(* Logix 5000 project; controller NWGG_Treater_Dayton vendor 1 type 14 code 238 rev 35.11; software revision 35.00; part 4 of 5 *)
(* tags used below, declared in another part *)
   Auto_Start_Treater : BOOL;
   Chemicals_Required : BOOL;
   Clear_Treater_Fault : BOOL;
   Current_Treater_Speed_Percent : REAL;
   Grain_Rate_CWT : REAL;
   IDX : DINT;
   K_Valve_ACK : BOOL;
   Manual_Start_Treater : BOOL;
   Non_Water_Total_Chemical_Package : REAL;
   Non_Water_Treatment_Package : REAL;
   SAIZeroScale : SAI_Zero_Scale[30];
   Start_Treating : BOOL;
   Stop_Treater : BOOL;
   tmrStartTreat : TIMER;
   tmrStopTreat : TIMER;
   Total_Chemical_Package : REAL;
   Treater_Pump : Treater_Pump[50];
   Treater_Running : BOOL;
   Treater_Speed_Percent : REAL;
   Water : Analog_Gallon_Values;
   Water_Control : Water_Pump_Control;
(* MainProgram, continued *)

ROUTINE Set_Scale_Values   (* ladder *)
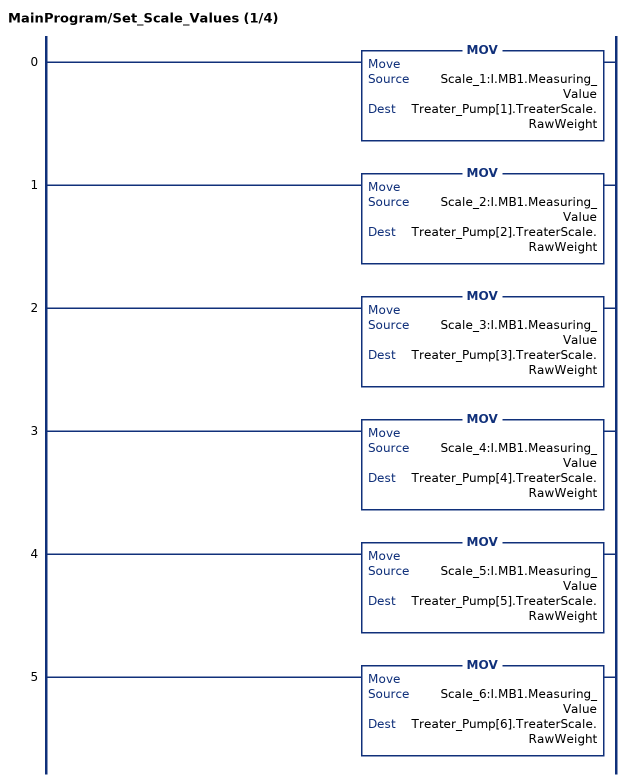
   0: MOV(Scale_1:I.MB1.Measuring_Value,Treater_Pump[1].TreaterScale.RawWeight);
   1: MOV(Scale_2:I.MB1.Measuring_Value,Treater_Pump[2].TreaterScale.RawWeight);
   2: MOV(Scale_3:I.MB1.Measuring_Value,Treater_Pump[3].TreaterScale.RawWeight);
   3: MOV(Scale_4:I.MB1.Measuring_Value,Treater_Pump[4].TreaterScale.RawWeight);
   4: MOV(Scale_5:I.MB1.Measuring_Value,Treater_Pump[5].TreaterScale.RawWeight);
   5: MOV(Scale_6:I.MB1.Measuring_Value,Treater_Pump[6].TreaterScale.RawWeight);
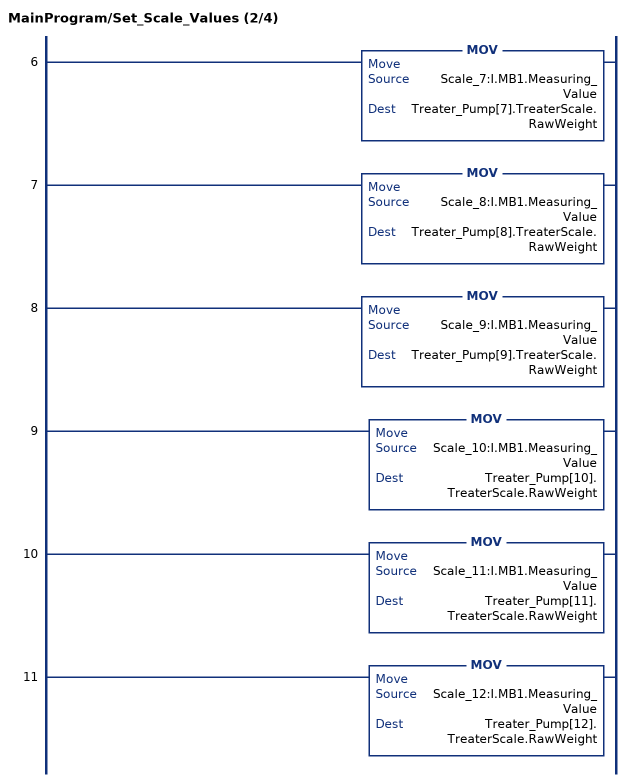
   6: MOV(Scale_7:I.MB1.Measuring_Value,Treater_Pump[7].TreaterScale.RawWeight);
   7: MOV(Scale_8:I.MB1.Measuring_Value,Treater_Pump[8].TreaterScale.RawWeight);
   8: MOV(Scale_9:I.MB1.Measuring_Value,Treater_Pump[9].TreaterScale.RawWeight);
   9: MOV(Scale_10:I.MB1.Measuring_Value,Treater_Pump[10].TreaterScale.RawWeight);
   10: MOV(Scale_11:I.MB1.Measuring_Value,Treater_Pump[11].TreaterScale.RawWeight);
   11: MOV(Scale_12:I.MB1.Measuring_Value,Treater_Pump[12].TreaterScale.RawWeight);
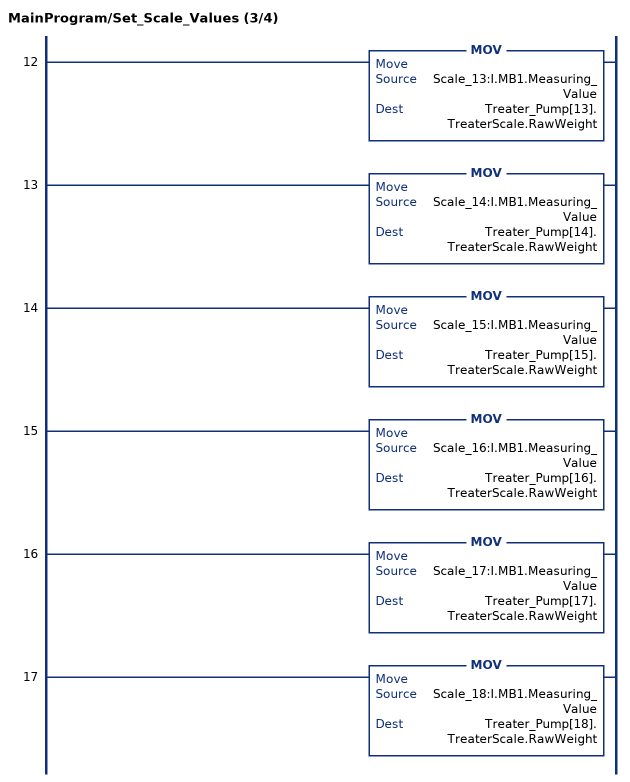
   12: MOV(Scale_13:I.MB1.Measuring_Value,Treater_Pump[13].TreaterScale.RawWeight);
   13: MOV(Scale_14:I.MB1.Measuring_Value,Treater_Pump[14].TreaterScale.RawWeight);
   14: MOV(Scale_15:I.MB1.Measuring_Value,Treater_Pump[15].TreaterScale.RawWeight);
   15: MOV(Scale_16:I.MB1.Measuring_Value,Treater_Pump[16].TreaterScale.RawWeight);
   16: MOV(Scale_17:I.MB1.Measuring_Value,Treater_Pump[17].TreaterScale.RawWeight);
   17: MOV(Scale_18:I.MB1.Measuring_Value,Treater_Pump[18].TreaterScale.RawWeight);
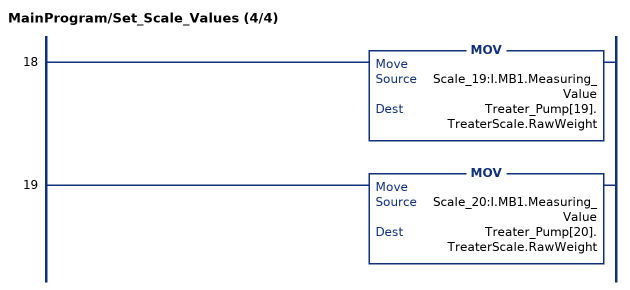
   18: MOV(Scale_19:I.MB1.Measuring_Value,Treater_Pump[19].TreaterScale.RawWeight);
   19: MOV(Scale_20:I.MB1.Measuring_Value,Treater_Pump[20].TreaterScale.RawWeight);
END_ROUTINE

ROUTINE SetHMIArrayIndex   (* ladder *)
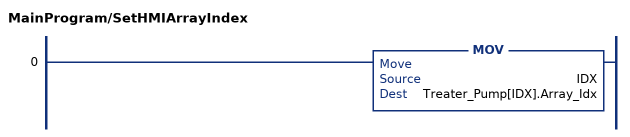
   0: MOV(IDX,Treater_Pump[IDX].Array_Idx);
END_ROUTINE

ROUTINE Treater   (* ladder *)
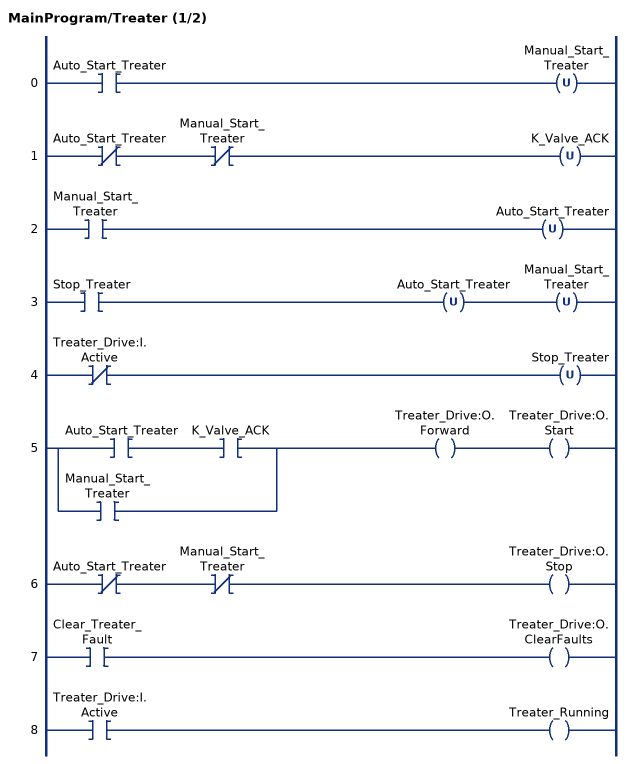
   0: XIC(Auto_Start_Treater)OTU(Manual_Start_Treater);
   1: XIO(Auto_Start_Treater)XIO(Manual_Start_Treater)OTU(K_Valve_ACK);
   2: XIC(Manual_Start_Treater)OTU(Auto_Start_Treater);
   3: XIC(Stop_Treater)OTU(Auto_Start_Treater)OTU(Manual_Start_Treater);
   4: XIO(Treater_Drive:I.Active)OTU(Stop_Treater);
   5: [XIC(Auto_Start_Treater) XIC(K_Valve_ACK) ,XIC(Manual_Start_Treater) ]OTE(Treater_Drive:O.Forward)OTE(Treater_Drive:O.Start);
   6: XIO(Auto_Start_Treater)XIO(Manual_Start_Treater)OTE(Treater_Drive:O.Stop);
   7: XIC(Clear_Treater_Fault)OTE(Treater_Drive:O.ClearFaults);
   8: XIC(Treater_Drive:I.Active)OTE(Treater_Running);
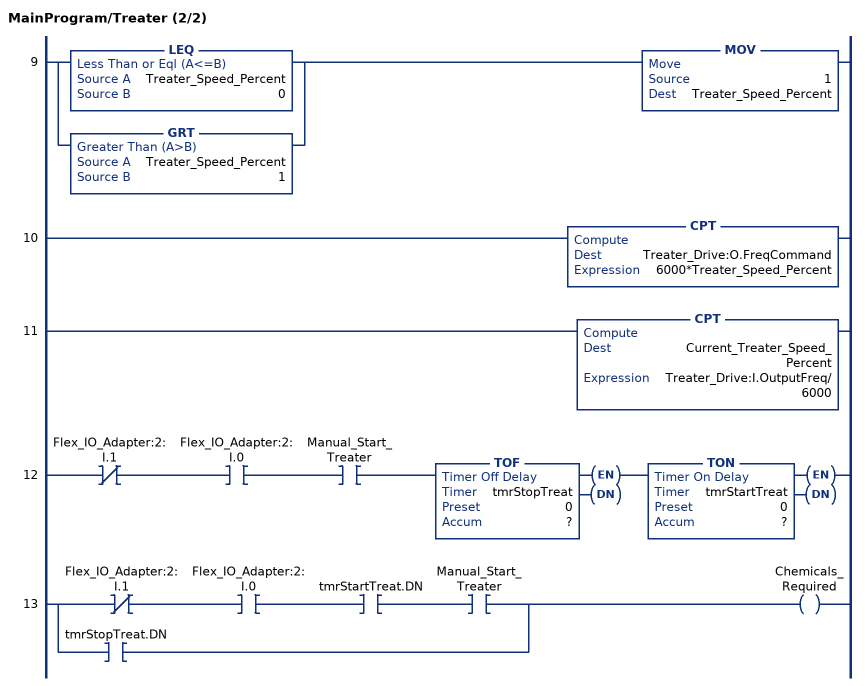
   9: [LEQ(Treater_Speed_Percent,0) ,GRT(Treater_Speed_Percent,1) ]MOV(1,Treater_Speed_Percent);
   10: CPT(Treater_Drive:O.FreqCommand,6000*Treater_Speed_Percent);
   11: CPT(Current_Treater_Speed_Percent,Treater_Drive:I.OutputFreq/6000);
   12: XIO(Flex_IO_Adapter:2:I.1)XIC(Flex_IO_Adapter:2:I.0)XIC(Manual_Start_Treater)TOF(tmrStopTreat,?,?)TON(tmrStartTreat,?,?);
   13: [XIO(Flex_IO_Adapter:2:I.1) XIC(Flex_IO_Adapter:2:I.0) XIC(tmrStartTreat.DN) XIC(Manual_Start_Treater) ,XIC(tmrStopTreat.DN) ]OTE(Chemicals_Required);
END_ROUTINE

ROUTINE Zero_Scales   (* ladder *)
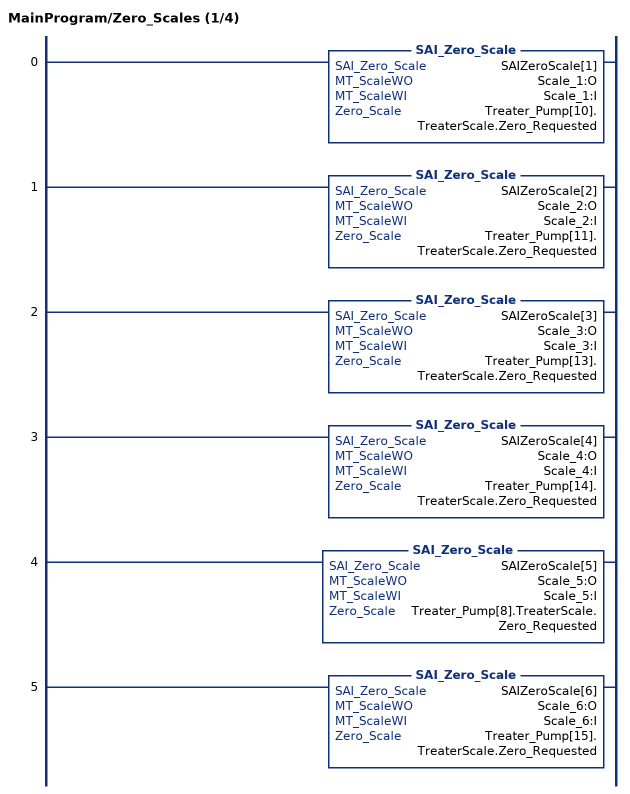
   0: SAI_Zero_Scale(SAIZeroScale[1],Scale_1:O,Scale_1:I,Treater_Pump[10].TreaterScale.Zero_Requested);
   1: SAI_Zero_Scale(SAIZeroScale[2],Scale_2:O,Scale_2:I,Treater_Pump[11].TreaterScale.Zero_Requested);
   2: SAI_Zero_Scale(SAIZeroScale[3],Scale_3:O,Scale_3:I,Treater_Pump[13].TreaterScale.Zero_Requested);
   3: SAI_Zero_Scale(SAIZeroScale[4],Scale_4:O,Scale_4:I,Treater_Pump[14].TreaterScale.Zero_Requested);
   4: SAI_Zero_Scale(SAIZeroScale[5],Scale_5:O,Scale_5:I,Treater_Pump[8].TreaterScale.Zero_Requested);
   5: SAI_Zero_Scale(SAIZeroScale[6],Scale_6:O,Scale_6:I,Treater_Pump[15].TreaterScale.Zero_Requested);
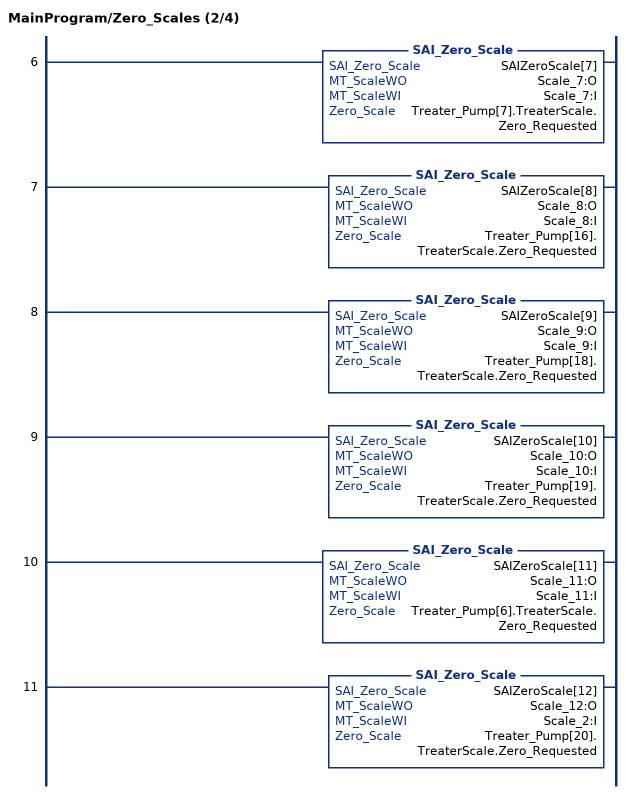
   6: SAI_Zero_Scale(SAIZeroScale[7],Scale_7:O,Scale_7:I,Treater_Pump[7].TreaterScale.Zero_Requested);
   7: SAI_Zero_Scale(SAIZeroScale[8],Scale_8:O,Scale_8:I,Treater_Pump[16].TreaterScale.Zero_Requested);
   8: SAI_Zero_Scale(SAIZeroScale[9],Scale_9:O,Scale_9:I,Treater_Pump[18].TreaterScale.Zero_Requested);
   9: SAI_Zero_Scale(SAIZeroScale[10],Scale_10:O,Scale_10:I,Treater_Pump[19].TreaterScale.Zero_Requested);
   10: SAI_Zero_Scale(SAIZeroScale[11],Scale_11:O,Scale_11:I,Treater_Pump[6].TreaterScale.Zero_Requested);
   11: SAI_Zero_Scale(SAIZeroScale[12],Scale_12:O,Scale_2:I,Treater_Pump[20].TreaterScale.Zero_Requested);
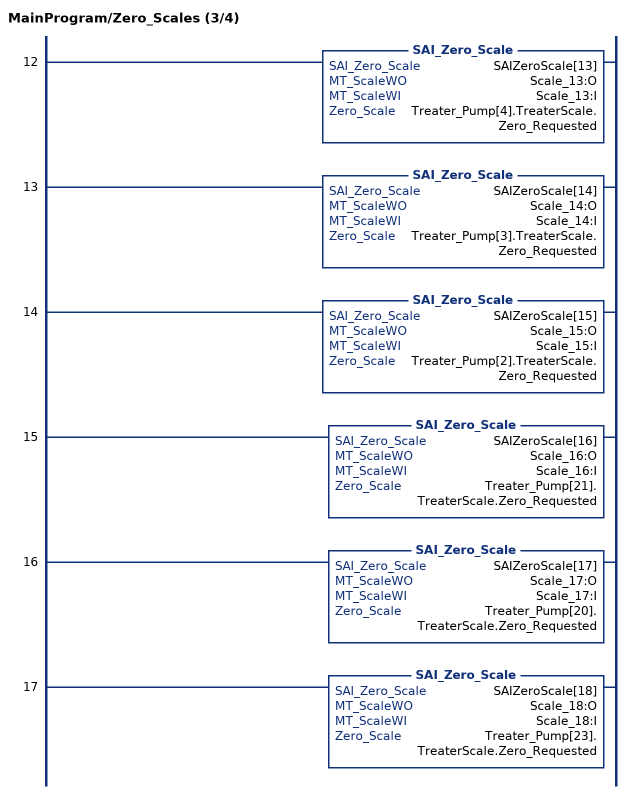
   12: SAI_Zero_Scale(SAIZeroScale[13],Scale_13:O,Scale_13:I,Treater_Pump[4].TreaterScale.Zero_Requested);
   13: SAI_Zero_Scale(SAIZeroScale[14],Scale_14:O,Scale_14:I,Treater_Pump[3].TreaterScale.Zero_Requested);
   14: SAI_Zero_Scale(SAIZeroScale[15],Scale_15:O,Scale_15:I,Treater_Pump[2].TreaterScale.Zero_Requested);
   15: SAI_Zero_Scale(SAIZeroScale[16],Scale_16:O,Scale_16:I,Treater_Pump[21].TreaterScale.Zero_Requested);
   16: SAI_Zero_Scale(SAIZeroScale[17],Scale_17:O,Scale_17:I,Treater_Pump[20].TreaterScale.Zero_Requested);
   17: SAI_Zero_Scale(SAIZeroScale[18],Scale_18:O,Scale_18:I,Treater_Pump[23].TreaterScale.Zero_Requested);
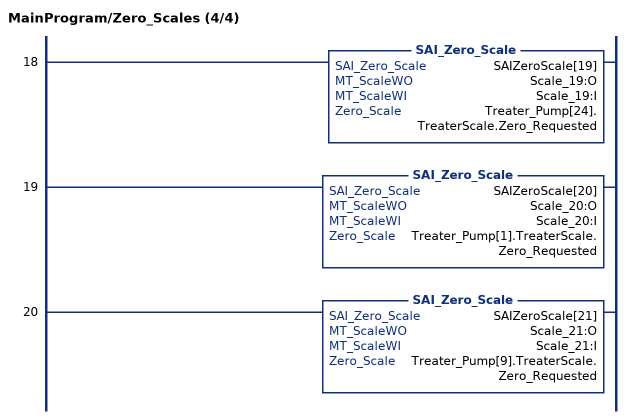
   18: SAI_Zero_Scale(SAIZeroScale[19],Scale_19:O,Scale_19:I,Treater_Pump[24].TreaterScale.Zero_Requested);
   19: SAI_Zero_Scale(SAIZeroScale[20],Scale_20:O,Scale_20:I,Treater_Pump[1].TreaterScale.Zero_Requested);
   20: SAI_Zero_Scale(SAIZeroScale[21],Scale_21:O,Scale_21:I,Treater_Pump[9].TreaterScale.Zero_Requested);
END_ROUTINE
END_PROGRAM

PROGRAM Pumps   (* main routine MainRoutine *)
VAR
   Active_Pump_Count_Changed : BOOL;
   Ant : BOOL;
   Auto_Start_Pumps : BOOL;
   Auto_Stop_Pumps : BOOL := 1;
   Calibrating_Pump : BOOL;
   Cancel_Cal : BOOL;
   Clear_All_Pump_Faults : BOOL;
   Current_Treatment_Count : DINT := 9;
   Default_Oil : DINT := 22;
   Default_Water : DINT := 220;   // The Default Water Per Min Used
   Manual_Water_Flush : BOOL;
   Prev_Treatment_Count : DINT := 9;
   Pump_Scale_Control : Pump_Scale_Control[50];
   Pumps_In_Fault : BOOL := 1;
   Reset_Treatments : BOOL;
   Start_Water_Flush : BOOL;
   Start_Water_Flush_ONS : BOOL := 1;
   tmrWaterFlush : TIMER;
   Water_Flush : BOOL;
END_VAR

ROUTINE Active_Treater_Pump_Count   (* ladder *)
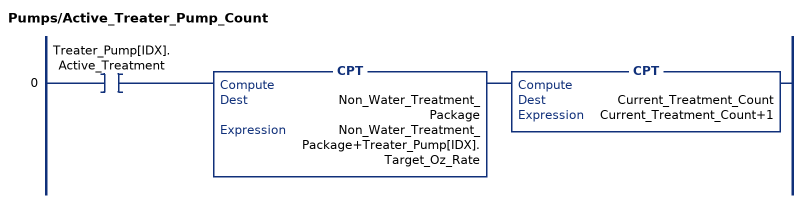
   0: XIC(Treater_Pump[IDX].Active_Treatment)CPT(Non_Water_Treatment_Package,Non_Water_Treatment_Package+Treater_Pump[IDX].Target_Oz_Rate)CPT(Current_Treatment_Count,Current_Treatment_Count+1);
END_ROUTINE

ROUTINE Check_Pump_Fault   (* ladder *)
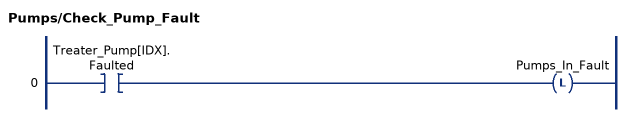
   0: XIC(Treater_Pump[IDX].Faulted)OTL(Pumps_In_Fault);
END_ROUTINE

ROUTINE Clear_All_Faults   (* ladder *)
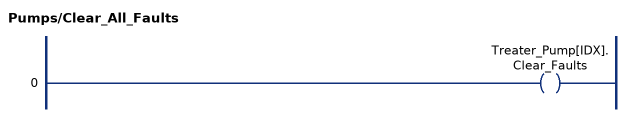
   0: OTE(Treater_Pump[IDX].Clear_Faults);
END_ROUTINE

ROUTINE MainRoutine   (* ladder *)
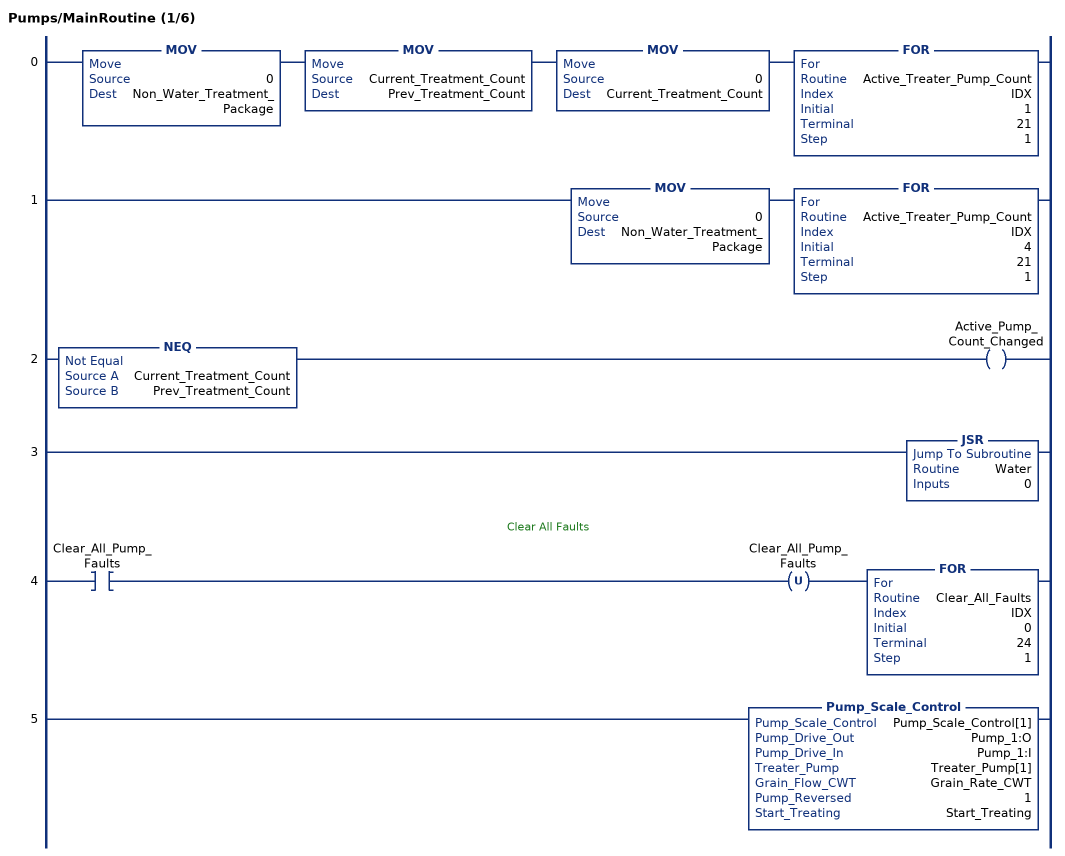
   0: MOV(0,Non_Water_Treatment_Package)MOV(Current_Treatment_Count,Prev_Treatment_Count)MOV(0,Current_Treatment_Count)FOR(Active_Treater_Pump_Count,IDX,1,21,1);
   1: MOV(0,Non_Water_Treatment_Package)FOR(Active_Treater_Pump_Count,IDX,4,21,1);
   2: NEQ(Current_Treatment_Count,Prev_Treatment_Count)OTE(Active_Pump_Count_Changed);
   3: JSR(Water,0);
   // Clear All Faults
   4: XIC(Clear_All_Pump_Faults)OTU(Clear_All_Pump_Faults)FOR(Clear_All_Faults,IDX,0,24,1);
   5: Pump_Scale_Control(Pump_Scale_Control[1],Pump_1:O,Pump_1:I,Treater_Pump[1],Grain_Rate_CWT,1,Start_Treating);
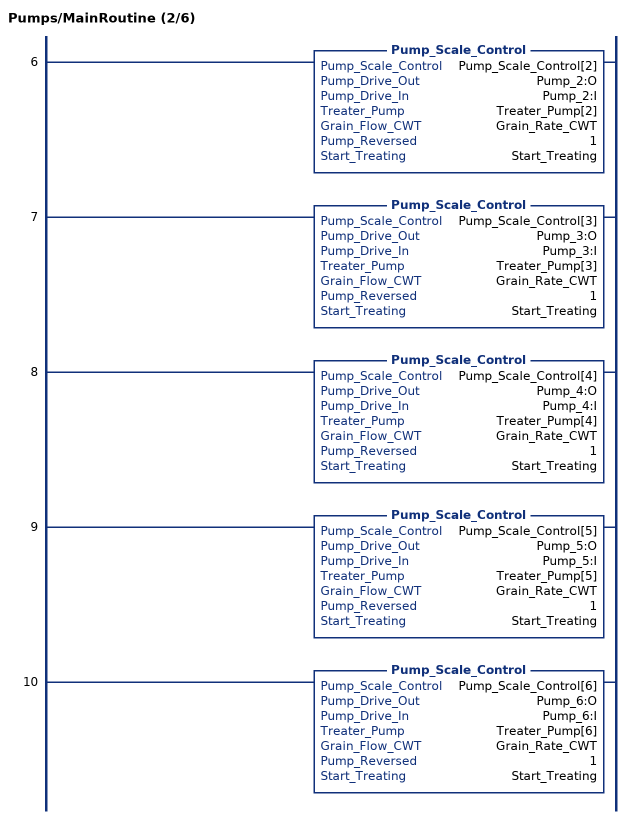
   6: Pump_Scale_Control(Pump_Scale_Control[2],Pump_2:O,Pump_2:I,Treater_Pump[2],Grain_Rate_CWT,1,Start_Treating);
   7: Pump_Scale_Control(Pump_Scale_Control[3],Pump_3:O,Pump_3:I,Treater_Pump[3],Grain_Rate_CWT,1,Start_Treating);
   8: Pump_Scale_Control(Pump_Scale_Control[4],Pump_4:O,Pump_4:I,Treater_Pump[4],Grain_Rate_CWT,1,Start_Treating);
   9: Pump_Scale_Control(Pump_Scale_Control[5],Pump_5:O,Pump_5:I,Treater_Pump[5],Grain_Rate_CWT,1,Start_Treating);
   10: Pump_Scale_Control(Pump_Scale_Control[6],Pump_6:O,Pump_6:I,Treater_Pump[6],Grain_Rate_CWT,1,Start_Treating);
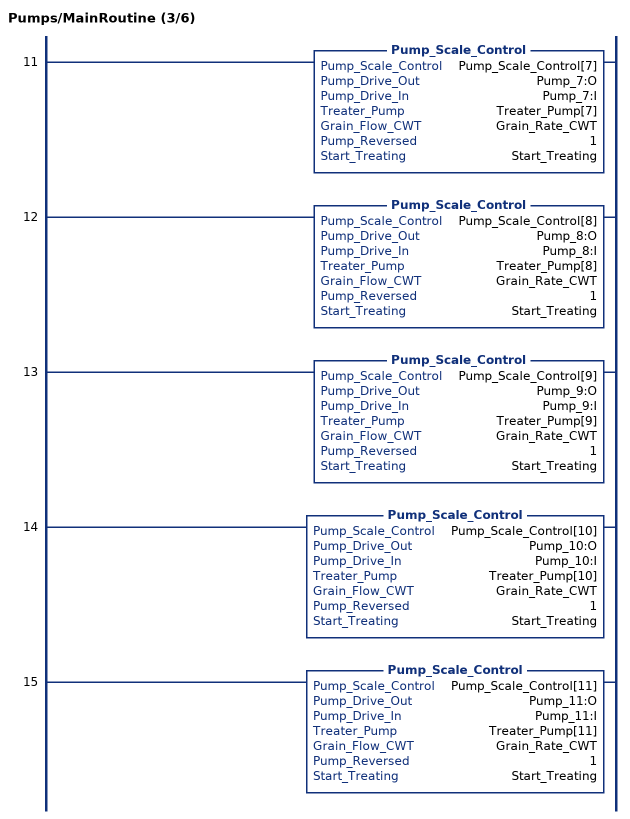
   11: Pump_Scale_Control(Pump_Scale_Control[7],Pump_7:O,Pump_7:I,Treater_Pump[7],Grain_Rate_CWT,1,Start_Treating);
   12: Pump_Scale_Control(Pump_Scale_Control[8],Pump_8:O,Pump_8:I,Treater_Pump[8],Grain_Rate_CWT,1,Start_Treating);
   13: Pump_Scale_Control(Pump_Scale_Control[9],Pump_9:O,Pump_9:I,Treater_Pump[9],Grain_Rate_CWT,1,Start_Treating);
   14: Pump_Scale_Control(Pump_Scale_Control[10],Pump_10:O,Pump_10:I,Treater_Pump[10],Grain_Rate_CWT,1,Start_Treating);
   15: Pump_Scale_Control(Pump_Scale_Control[11],Pump_11:O,Pump_11:I,Treater_Pump[11],Grain_Rate_CWT,1,Start_Treating);
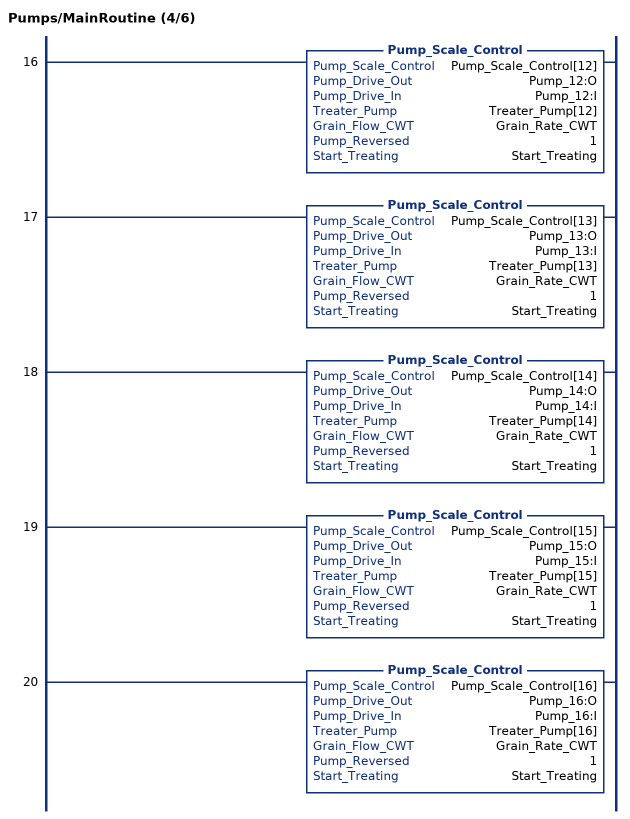
   16: Pump_Scale_Control(Pump_Scale_Control[12],Pump_12:O,Pump_12:I,Treater_Pump[12],Grain_Rate_CWT,1,Start_Treating);
   17: Pump_Scale_Control(Pump_Scale_Control[13],Pump_13:O,Pump_13:I,Treater_Pump[13],Grain_Rate_CWT,1,Start_Treating);
   18: Pump_Scale_Control(Pump_Scale_Control[14],Pump_14:O,Pump_14:I,Treater_Pump[14],Grain_Rate_CWT,1,Start_Treating);
   19: Pump_Scale_Control(Pump_Scale_Control[15],Pump_15:O,Pump_15:I,Treater_Pump[15],Grain_Rate_CWT,1,Start_Treating);
   20: Pump_Scale_Control(Pump_Scale_Control[16],Pump_16:O,Pump_16:I,Treater_Pump[16],Grain_Rate_CWT,1,Start_Treating);
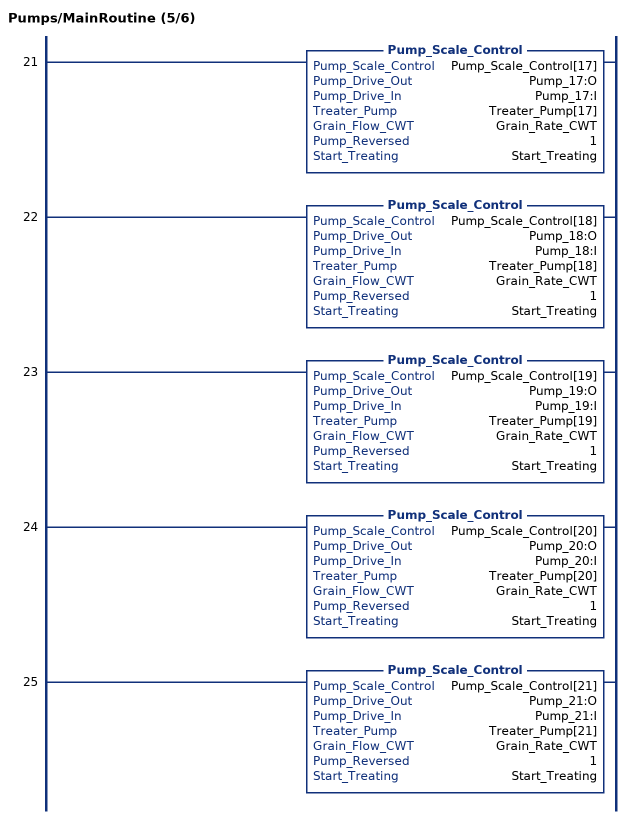
   21: Pump_Scale_Control(Pump_Scale_Control[17],Pump_17:O,Pump_17:I,Treater_Pump[17],Grain_Rate_CWT,1,Start_Treating);
   22: Pump_Scale_Control(Pump_Scale_Control[18],Pump_18:O,Pump_18:I,Treater_Pump[18],Grain_Rate_CWT,1,Start_Treating);
   23: Pump_Scale_Control(Pump_Scale_Control[19],Pump_19:O,Pump_19:I,Treater_Pump[19],Grain_Rate_CWT,1,Start_Treating);
   24: Pump_Scale_Control(Pump_Scale_Control[20],Pump_20:O,Pump_20:I,Treater_Pump[20],Grain_Rate_CWT,1,Start_Treating);
   25: Pump_Scale_Control(Pump_Scale_Control[21],Pump_21:O,Pump_21:I,Treater_Pump[21],Grain_Rate_CWT,1,Start_Treating);
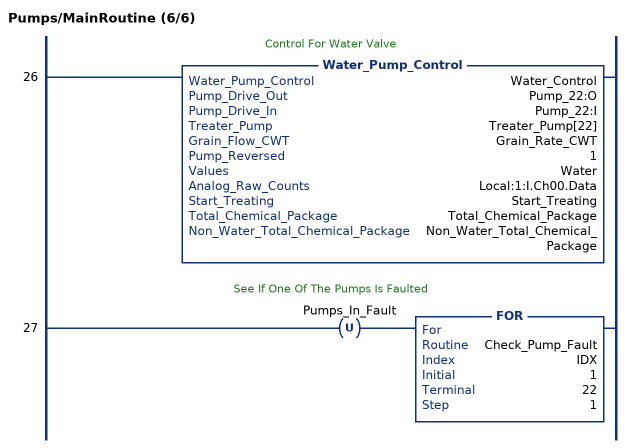
   // Control For Water Valve
   26: Water_Pump_Control(Water_Control,Pump_22:O,Pump_22:I,Treater_Pump[22],Grain_Rate_CWT,1,Water,Local:1:I.Ch00.Data,Start_Treating,Total_Chemical_Package,Non_Water_Total_Chemical_Package);
   // See If One Of The Pumps Is Faulted
   27: OTU(Pumps_In_Fault)FOR(Check_Pump_Fault,IDX,1,22,1);
END_ROUTINE
